DATA_BLOCK "db3006i_BC56_BancoCarga"
TITLE = db3006i_BC56_BancoCarga (DB3006)
AUTHOR : 'RegLobo'
VERSION : 0.1
////====================================
//// DB de INSTANCIA ("i" no nome = instancia, padrao do projeto) do fb_bancoCarga16 para o banco BC56. Numero DB3006 (base 3000 + 6). Importe DEPOIS do fb_bancoCarga16 e ANTES do fc_bancosCarga1200.
//// (o outro DB do banco e o de TELEGRAMA, db3007_BC56_Com, em db_ComBancos.) Se o TIA numerar diferente, ajuste o numero nas propriedades do bloco (numeracao manual).
////====================================
"fb_bancoCarga16"
BEGIN
END_DATA_BLOCK
